PROGRAM main
  VAR
    S1 AT %IX0.0 : BOOL; (* pulsador NA *)
    S2 AT %IX0.1 : BOOL; (* pulsador NA *)
    H1 AT %QX0.0 : BOOL; (* piloto verde *)
    H2 AT %QX0.1 : BOOL; (* piloto amarillo *)
  END_VAR
  VAR  (* added by the conversion: wires and edge detectors of the diagram *)
    _NOT1_OUT : BOOL;
  END_VAR

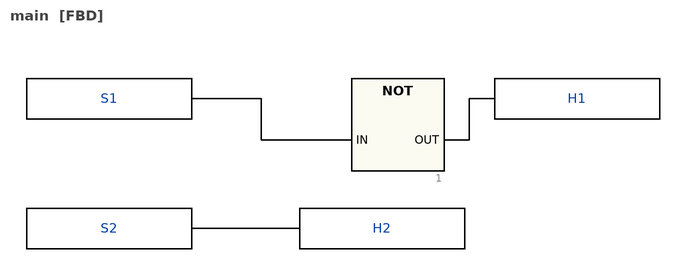
(* FBD diagram, written out as Structured Text *)
_NOT1_OUT := NOT S1;
H1 := _NOT1_OUT;
H2 := S2;
END_PROGRAM
